Fanuc KAREL source: KT00840.KL

PROGRAM KT00840
%NOLOCKGROUP
VAR
  B1: BOOLEAN
  B2: BOOLEAN
  OUT: INTEGER
BEGIN
  B1 = TRUE
  B2 = FALSE
  B1 = TRUE
  B2 = FALSE
  OUT = SQRT(B1)
END KT00840
